Fanuc KAREL source: KA00042.KL

PROGRAM KA00042
%NOLOCKGROUP
VAR
  SRC: STRING[80]
  DST: XYZWPR
BEGIN
  SRC = 'A'
  DST = SRC
END KA00042
